(* IEC 61131-3 sources: brew/plc/plc-cellar, 2 files *)

(* ---- plc-cellar-plant.st ---- *)
(*
  plc-cellar: CherryMountain Brewery cellar PLC, full and lite variants
  (DESIGN.md 6.3, 6.7, 12.1). The ci slice runs plc-cellar.st instead.

  Per fermenter FV-101 .. FV-104:
    - on/off glycol valve control with a 0.5 degF hysteresis half band on the
      side and cone zones (cooling only)
    - the spunding setpoint: 1 psig while the beer is fermenting, 12 psig once
      the apparent extract falls below 5 degP (near terminal gravity), written
      to the RIO as absolute pressure every scan
    - the fermentation profile (FermentProfile): while CEL.PROFILE.HSnn.AUTO is
      set, the program writes both temperature setpoints for the beer's stage,
      66 degF fermenting, 70 degF for the diacetyl rest, 34 degF for the crash
      (CEL.PROFILE.TC01 to TC03, the operator's), and shows the stage in
      KSnn.STAGE. The rest lasts KC01 minutes: 180, which is 144 h of
      fermentation on the range's 48x clock. With AUTO clear the setpoints are
      the operator's. A crash raises the fermenter's temperature deviation
      alarms until the beer is cold.
  Per bright tank BBT-201 and BBT-202:
    - jacket glycol valve on/off control
    - the equilibrium head pressure for the carbonation target at the
      temperature setpoint (Zahm-Nagel fit, sea-level gauge plus 14.7 psi =
      absolute; the setpoint, not the measured temperature, so the limit does
      not swing with the glycol hysteresis), and carbonation-stone flow
      proportional to the shortfall in dissolved CO2, closed while the head is
      more than HEAD_MARGIN above that pressure or at HEAD_MAX (0.5 psi under
      the 26.1 psia high-pressure alarm), so neither that alarm nor the 15 psig
      relief valve trips in normal running. A target whose equilibrium is above
      HEAD_MAX - HEAD_MARGIN cannot be reached, so AT01.SP is clamped to the
      most that can (VOL_MAX, solved from the same fit), and the HMI shows it.
    - BBT-202 feeds the bottling line: its outlet opens while it holds beer
  Shared equipment:
    - the cellar CO2 life-safety interlock (DESIGN.md 6.7): CEL.SYS.XS01.CO2_OK
      is the hardwired, de-energize-to-trip relay from bas-vent. While it is
      open, and for CO2_RELEASE_DELAY after it closes again, the program sets
      CO2_INHIBIT, closes both carbonation valves, and closes the hop-port CO2
      purge (holding a dry-hop sequence in its purge step). No supervisory host
      takes part. The relay reads open until the building federate first
      reports it, so carbonation starts inhibited.
    - the dry-hop sequence on an operator request: CO2 purge, then dose
    - the transfer and CIP peer status bits that plc-utilities reads
    - confined-space entry (29 CFR 1910.146, DESIGN.md 6.3): a vessel's entry
      permit bit locks out its glycol valves, the bright tanks' carbonation
      stone and outlet, and (through plc-utilities) its CIP circuit, vents a
      fermenter's head through its spunding valve, holds the dry-hop doser
      while any fermenter is entered, and latches a critical alarm when a
      locked-out output is found written between scans
  Alarms (every bit in alarms.json for this PLC) are generated by
  plc/common/plcbuild.py at the ALARMS marker, with their deadbands and delays.

  Units: analog values are raw registers, engineering value x 10^scaling
  (degF x 100, psia x 100, vol x 100, % x 10). Setpoints in %MW belong to the
  operator after the first scan; the program loads defaults once and clamps.
*)

(* One glycol zone: cooling-only on/off valve with hysteresis. *)
FUNCTION_BLOCK GlycolZone
  VAR_INPUT
    PV : UINT;                 (* temperature, degF x 100 *)
    SP : UINT;                 (* setpoint, degF x 100 *)
    HYST : UINT := 50;         (* half band, 0.5 degF *)
  END_VAR
  VAR_OUTPUT
    VALVE : BOOL;              (* TRUE = open (cooling) *)
  END_VAR
  IF PV >= SP + HYST THEN
    VALVE := TRUE;
  ELSIF PV + HYST <= SP THEN
    VALVE := FALSE;
  END_IF;
END_FUNCTION_BLOCK

(* Carbonation for one bright tank. *)
FUNCTION_BLOCK Carbonation
  VAR_INPUT
    TEMP_SP : UINT;            (* temperature setpoint, degF x 100 *)
    VOL_SP : UINT;             (* target, vol x 100 *)
    VOL_PV : UINT;             (* inline meter, vol x 100 *)
    PSIA_PV : UINT;            (* head pressure, psia x 100 *)
    INHIBIT : BOOL;            (* cellar CO2 interlock *)
    HEAD_MARGIN : UINT := 50;  (* stone closes 0.5 psi above equilibrium, psi x 100 *)
    HEAD_MAX : UINT := 2560;   (* and never above 25.6 psia, psia x 100 *)
  END_VAR
  VAR_OUTPUT
    PSIA_SP : UINT;            (* equilibrium head pressure, psia x 100 *)
    VALVE : UINT;              (* stone flow valve, % x 10 *)
    VOL_MAX : UINT;            (* most reachable under HEAD_MAX, vol x 100 *)
  END_VAR
  VAR
    temp_f : REAL;
    vol : REAL;
    psig_sea_level : REAL;
    shortfall : REAL;
    qa : REAL;
    qb : REAL;
    qc : REAL;
  END_VAR
  temp_f := UINT_TO_REAL(TEMP_SP) / 100.0;
  (* The fit is quadratic in vol: qa vol^2 + qb vol + qc = 0 at the highest
     equilibrium the stone may build to (HEAD_MAX - HEAD_MARGIN). *)
  qa := -0.0684226;
  qb := 4.24267 + 0.173354 * temp_f;
  qc := -16.6999 - 0.0101059 * temp_f + 0.00116512 * temp_f * temp_f
    - (UINT_TO_REAL(HEAD_MAX - HEAD_MARGIN) / 100.0 - 14.7);
  VOL_MAX := REAL_TO_UINT(LIMIT(0.0,
    (SQRT(qb * qb - 4.0 * qa * qc) - qb) / (2.0 * qa) * 100.0, 500.0));
  vol := UINT_TO_REAL(MIN(VOL_SP, VOL_MAX)) / 100.0;
  psig_sea_level := -16.6999 - 0.0101059 * temp_f + 0.00116512 * temp_f * temp_f
    + 0.173354 * temp_f * vol + 4.24267 * vol - 0.0684226 * vol * vol;
  PSIA_SP := REAL_TO_UINT(LIMIT(0.0, (psig_sea_level + 14.7) * 100.0, 4000.0));
  (* 100 % at 0.5 vol or more short of the target, closed at the target. *)
  shortfall := vol - UINT_TO_REAL(VOL_PV) / 100.0;
  IF INHIBIT OR shortfall <= 0.0 OR PSIA_PV >= MIN(PSIA_SP + HEAD_MARGIN, HEAD_MAX) THEN
    VALVE := 0;
  ELSE
    VALVE := REAL_TO_UINT(LIMIT(0.0, shortfall * 2000.0, 1000.0));
  END_IF;
END_FUNCTION_BLOCK

(* The fermentation profile of one fermenter (DESIGN.md 6.3): which stage the
   beer is in, and the temperature that goes with it. A stage follows from the
   density meter: a vessel that reads no extract is empty, wort above TERMINAL is
   fermenting, and beer under it rests warm for REST_MIN minutes (counted in
   scans) and is then crashed. A reading must hold for SETTLE_MS before it ends
   a stage: a meter that drops out for a scan or a few seconds has not emptied
   the vessel or finished the fermentation, and the stage it would end is one
   the program cannot get back to. Beer the program has not followed from its
   fill (after a start of the PLC) is taken as crashed when it is already cold,
   and as starting its rest otherwise.

   The setpoint is one the vessel can follow, so that the deviation alarm means
   a fault and not a stage:
   - A fermenter has jackets and no heater. On the way up (wort pitched under
     the fermentation temperature, the free rise to the rest) the setpoint
     leads the beer by LEAD and goes no higher than the stage's temperature. It
     does not come back down with the beer: beer that cools in these stages has
     a glycol valve that leaks. Only a fill is different: for FILL_MS after a
     fermentation starts the setpoint follows the vessel down too, to the
     temperature of the wort that is coming in.
   - The crash falls from where the beer is toward the glycol's temperature, by
     CRASH_PCT_H percent of what is left each hour, and stops at CRASH_SP. That
     is the curve of a jacketed tank, a little slower than this one cools, so
     beer that falls behind it has lost its cooling.
   - An empty vessel's setpoint stays LEAD above the vessel: its jackets stay
     shut, the next wort is not chilled on its way in, and nothing alarms. *)
FUNCTION_BLOCK FermentProfile
  VAR_INPUT
    EXTRACT : UINT;            (* apparent extract, degP x 100 *)
    TEMP : UINT;               (* side temperature, degF x 100 *)
    FERMENT_SP : UINT;         (* temperature while fermenting, degF x 100 *)
    REST_SP : UINT;            (* temperature of the diacetyl rest, degF x 100 *)
    CRASH_SP : UINT;           (* temperature of the crash, degF x 100 *)
    REST_MIN : UINT;           (* rest length, minutes *)
    SCAN_MS : UDINT;           (* the task interval, ms *)
    EMPTY : UINT := 50;        (* under 0.5 degP the vessel is empty *)
    TERMINAL : UINT := 500;    (* under 5 degP the beer is near terminal gravity *)
    COLD : UINT := 6000;       (* under 60 degF the beer has been crashed *)
    SETTLE_MS : UDINT := 60000;  (* a reading ends a stage once it has held this long *)
    LEAD : UINT := 100;        (* on the way up the setpoint leads the beer by 1 degF *)
    GLYCOL : UINT := 2800;     (* the glycol supply, degF x 100: the crash falls toward it *)
    CRASH_PCT_H : UINT := 25;  (* ... by this share of what is left, each hour *)
    SP_MIN : UINT := 2000;     (* the setpoint limits of the program *)
    SP_MAX : UINT := 9000;
    FILL_MS : UDINT := 1800000;  (* a knockout into the vessel is over in this time *)
  END_VAR
  VAR_OUTPUT
    STAGE : UINT;              (* 0 empty, 1 fermenting, 2 diacetyl rest, 3 crash *)
    SP : UINT;                 (* the stage's setpoint now, degF x 100 *)
  END_VAR
  VAR
    rest_ms : UDINT;           (* time in the rest so far *)
    empty_ms : UDINT;          (* how long the meter has read no extract *)
    terminal_ms : UDINT;       (* how long it has read under TERMINAL *)
    last_stage : UINT := 99;   (* the stage of the scan before; 99 before the first *)
    sp_now : REAL := 0.0;      (* the setpoint, degF x 100, between scans *)
    lead_sp : REAL;
    cap : REAL;
    stage_ms : UDINT;          (* time in the stage, up to FILL_MS *)
  END_VAR
  IF EXTRACT < EMPTY THEN
    empty_ms := MIN(empty_ms + SCAN_MS, SETTLE_MS);
  ELSE
    empty_ms := 0;
  END_IF;
  IF EXTRACT < TERMINAL THEN
    terminal_ms := MIN(terminal_ms + SCAN_MS, SETTLE_MS);
  ELSE
    terminal_ms := 0;
  END_IF;
  IF EXTRACT < EMPTY THEN
    (* Until the reading has held, the stage stays as it is (and a rest's clock
       waits): this may be the meter, not the vessel. *)
    IF empty_ms >= SETTLE_MS THEN
      STAGE := 0;
    END_IF;
  ELSIF STAGE = 0 THEN
    IF EXTRACT >= TERMINAL THEN
      STAGE := 1;
    ELSIF TEMP < COLD THEN
      STAGE := 3;
    ELSE
      STAGE := 2;
      rest_ms := 0;
    END_IF;
  ELSIF STAGE = 1 THEN
    IF terminal_ms >= SETTLE_MS THEN
      STAGE := 2;
      rest_ms := 0;
    END_IF;
  ELSIF STAGE = 2 THEN
    IF rest_ms >= UINT_TO_UDINT(REST_MIN) * 60000 THEN
      STAGE := 3;
    ELSE
      rest_ms := rest_ms + SCAN_MS;
    END_IF;
  END_IF;

  lead_sp := UINT_TO_REAL(TEMP) + UINT_TO_REAL(LEAD);
  IF STAGE = 3 THEN
    IF last_stage <> 3 THEN
      sp_now := UINT_TO_REAL(TEMP);   (* the crash starts from where the beer is *)
    END_IF;
    sp_now := sp_now - (sp_now - UINT_TO_REAL(GLYCOL)) * UINT_TO_REAL(CRASH_PCT_H) / 100.0
      * UDINT_TO_REAL(SCAN_MS) / 3600000.0;
    sp_now := MAX(sp_now, UINT_TO_REAL(CRASH_SP));
  ELSIF STAGE = 0 THEN
    sp_now := lead_sp;
  ELSE
    IF STAGE = 2 THEN
      cap := UINT_TO_REAL(REST_SP);
    ELSE
      cap := UINT_TO_REAL(FERMENT_SP);
    END_IF;
    IF last_stage <> STAGE THEN
      stage_ms := 0;
      IF last_stage <> 1 THEN
        sp_now := 0.0;                (* nothing to carry over: start from the beer *)
      END_IF;
    ELSE
      stage_ms := MIN(stage_ms + SCAN_MS, FILL_MS);
    END_IF;
    IF STAGE = 1 AND stage_ms < FILL_MS THEN
      sp_now := MIN(cap, lead_sp);    (* a fill: down to the wort's temperature too *)
    ELSE
      sp_now := MIN(cap, MAX(sp_now, lead_sp));
    END_IF;
  END_IF;
  last_stage := STAGE;
  SP := REAL_TO_UINT(LIMIT(UINT_TO_REAL(SP_MIN), sp_now, UINT_TO_REAL(SP_MAX)));
END_FUNCTION_BLOCK

PROGRAM plc_cellar
  (* LOCATED_VARS: plcbuild.py splices the located variables and alarm instances here. *)

  VAR CONSTANT
    TEMP_SP_MIN : UINT := 2000;       (* 20 degF *)
    TEMP_SP_MAX : UINT := 9000;       (* 90 degF *)
    VOL_SP_MAX : UINT := 350;         (* 3.5 vol *)
    AMBIENT_PSIA : UINT := 1210;      (* 12.1 psia at 5,200 ft *)
    SPUND_LOW_PSIG : UINT := 100;     (* 1 psig while fermenting *)
    SPUND_HIGH_PSIG : UINT := 1200;   (* 12 psig near terminal gravity *)
    TERMINAL_PLATO : UINT := 500;     (* 5 degP *)
    BBT_FEED_MIN_LEVEL : UINT := 50;  (* 5 % *)
    CO2_RELEASE_DELAY : TIME := T#60s;  (* relay must be healthy this long *)
    DH_PURGE_TIME : TIME := T#30s;      (* hop-port CO2 purge before a dose *)
    DH_DOSE_TIME : TIME := T#60s;       (* dose valve open *)
    SCAN_MS : UDINT := 100;           (* the task interval plcbuild.py sets (T#100ms) *)
    REST_MIN_MAX : UINT := 6000;      (* 100 h *)
  END_VAR

  VAR
    started : BOOL := FALSE;
    fv101_side : GlycolZone;
    fv101_cone : GlycolZone;
    fv102_side : GlycolZone;
    fv102_cone : GlycolZone;
    fv103_side : GlycolZone;
    fv103_cone : GlycolZone;
    fv104_side : GlycolZone;
    fv104_cone : GlycolZone;
    fv101_profile : FermentProfile;
    fv102_profile : FermentProfile;
    fv103_profile : FermentProfile;
    fv104_profile : FermentProfile;
    bbt201_zone : GlycolZone;
    bbt202_zone : GlycolZone;
    bbt201_carb : Carbonation;
    bbt202_carb : Carbonation;
    co2_healthy : TON;
    transfer_active : BOOL;
    dh_step : INT := 0;
    dh_purge : TON;
    dh_dose : TON;
    fv_entry : BOOL;
  END_VAR

  (* First scan: default setpoints for the staggered initial state (DESIGN.md 9.4). *)
  IF NOT started THEN
    CEL_FV101_TT01_SP := 6600;
    CEL_FV101_TT02_SP := 6600;
    CEL_FV102_TT01_SP := 6600;
    CEL_FV102_TT02_SP := 6600;
    CEL_FV103_TT01_SP := 6800;
    CEL_FV103_TT02_SP := 6800;
    CEL_FV104_TT01_SP := 3400;
    CEL_FV104_TT02_SP := 3400;
    CEL_BBT201_TT01_SP := 3400;
    CEL_BBT202_TT01_SP := 3400;
    CEL_BBT201_AT01_SP := 260;
    CEL_BBT202_AT01_SP := 260;
    (* The recipe's profile (fire-of-the-phenix), on for every fermenter. *)
    CEL_PROFILE_TC01_SP := 6600;
    CEL_PROFILE_TC02_SP := 7000;
    CEL_PROFILE_TC03_SP := 3400;
    CEL_PROFILE_KC01_SP := 180;
    CEL_PROFILE_HS01_AUTO := TRUE;
    CEL_PROFILE_HS02_AUTO := TRUE;
    CEL_PROFILE_HS03_AUTO := TRUE;
    CEL_PROFILE_HS04_AUTO := TRUE;
    started := TRUE;
  END_IF;

  CEL_FV101_TT01_SP := LIMIT(TEMP_SP_MIN, CEL_FV101_TT01_SP, TEMP_SP_MAX);
  CEL_FV101_TT02_SP := LIMIT(TEMP_SP_MIN, CEL_FV101_TT02_SP, TEMP_SP_MAX);
  CEL_FV102_TT01_SP := LIMIT(TEMP_SP_MIN, CEL_FV102_TT01_SP, TEMP_SP_MAX);
  CEL_FV102_TT02_SP := LIMIT(TEMP_SP_MIN, CEL_FV102_TT02_SP, TEMP_SP_MAX);
  CEL_FV103_TT01_SP := LIMIT(TEMP_SP_MIN, CEL_FV103_TT01_SP, TEMP_SP_MAX);
  CEL_FV103_TT02_SP := LIMIT(TEMP_SP_MIN, CEL_FV103_TT02_SP, TEMP_SP_MAX);
  CEL_FV104_TT01_SP := LIMIT(TEMP_SP_MIN, CEL_FV104_TT01_SP, TEMP_SP_MAX);
  CEL_FV104_TT02_SP := LIMIT(TEMP_SP_MIN, CEL_FV104_TT02_SP, TEMP_SP_MAX);
  CEL_BBT201_TT01_SP := LIMIT(TEMP_SP_MIN, CEL_BBT201_TT01_SP, TEMP_SP_MAX);
  CEL_BBT202_TT01_SP := LIMIT(TEMP_SP_MIN, CEL_BBT202_TT01_SP, TEMP_SP_MAX);
  CEL_BBT201_AT01_SP := MIN(CEL_BBT201_AT01_SP, VOL_SP_MAX);
  CEL_BBT202_AT01_SP := MIN(CEL_BBT202_AT01_SP, VOL_SP_MAX);
  CEL_PROFILE_TC01_SP := LIMIT(TEMP_SP_MIN, CEL_PROFILE_TC01_SP, TEMP_SP_MAX);
  CEL_PROFILE_TC02_SP := LIMIT(TEMP_SP_MIN, CEL_PROFILE_TC02_SP, TEMP_SP_MAX);
  CEL_PROFILE_TC03_SP := LIMIT(TEMP_SP_MIN, CEL_PROFILE_TC03_SP, TEMP_SP_MAX);
  CEL_PROFILE_KC01_SP := MIN(CEL_PROFILE_KC01_SP, REST_MIN_MAX);

  (* ---- fermentation profile: the stage's temperature for a fermenter on AUTO --- *)
  fv101_profile(EXTRACT := CEL_FV101_DT01_PV, TEMP := CEL_FV101_TT01_PV,
    FERMENT_SP := CEL_PROFILE_TC01_SP, REST_SP := CEL_PROFILE_TC02_SP,
    CRASH_SP := CEL_PROFILE_TC03_SP, REST_MIN := CEL_PROFILE_KC01_SP, SCAN_MS := SCAN_MS);
  CEL_PROFILE_KS01_STAGE := fv101_profile.STAGE;
  IF CEL_PROFILE_HS01_AUTO THEN
    CEL_FV101_TT01_SP := fv101_profile.SP;
    CEL_FV101_TT02_SP := fv101_profile.SP;
  END_IF;
  fv102_profile(EXTRACT := CEL_FV102_DT01_PV, TEMP := CEL_FV102_TT01_PV,
    FERMENT_SP := CEL_PROFILE_TC01_SP, REST_SP := CEL_PROFILE_TC02_SP,
    CRASH_SP := CEL_PROFILE_TC03_SP, REST_MIN := CEL_PROFILE_KC01_SP, SCAN_MS := SCAN_MS);
  CEL_PROFILE_KS02_STAGE := fv102_profile.STAGE;
  IF CEL_PROFILE_HS02_AUTO THEN
    CEL_FV102_TT01_SP := fv102_profile.SP;
    CEL_FV102_TT02_SP := fv102_profile.SP;
  END_IF;
  fv103_profile(EXTRACT := CEL_FV103_DT01_PV, TEMP := CEL_FV103_TT01_PV,
    FERMENT_SP := CEL_PROFILE_TC01_SP, REST_SP := CEL_PROFILE_TC02_SP,
    CRASH_SP := CEL_PROFILE_TC03_SP, REST_MIN := CEL_PROFILE_KC01_SP, SCAN_MS := SCAN_MS);
  CEL_PROFILE_KS03_STAGE := fv103_profile.STAGE;
  IF CEL_PROFILE_HS03_AUTO THEN
    CEL_FV103_TT01_SP := fv103_profile.SP;
    CEL_FV103_TT02_SP := fv103_profile.SP;
  END_IF;
  fv104_profile(EXTRACT := CEL_FV104_DT01_PV, TEMP := CEL_FV104_TT01_PV,
    FERMENT_SP := CEL_PROFILE_TC01_SP, REST_SP := CEL_PROFILE_TC02_SP,
    CRASH_SP := CEL_PROFILE_TC03_SP, REST_MIN := CEL_PROFILE_KC01_SP, SCAN_MS := SCAN_MS);
  CEL_PROFILE_KS04_STAGE := fv104_profile.STAGE;
  IF CEL_PROFILE_HS04_AUTO THEN
    CEL_FV104_TT01_SP := fv104_profile.SP;
    CEL_FV104_TT02_SP := fv104_profile.SP;
  END_IF;

  (* ---- confined-space entry (29 CFR 1910.146, DESIGN.md 6.3) ------------------ *)
  (* The entry supervisor sets HSnn.ENTRY when the permit is issued. The program
     leaves every locked-out output off at the end of a scan, so a locked output
     that is on at the top of this one was written in between (an HMI, the EWS,
     or an attacker on the PLC's Modbus server): XAnn latches until the entry
     ends. *)
  CEL_ENTRY_XA01_PV := CEL_ENTRY_XS01_LOCKED
    AND (CEL_ENTRY_XA01_PV OR CEL_FV101_TV01_CMD OR CEL_FV101_TV02_CMD);
  CEL_ENTRY_XA02_PV := CEL_ENTRY_XS02_LOCKED
    AND (CEL_ENTRY_XA02_PV OR CEL_FV102_TV01_CMD OR CEL_FV102_TV02_CMD);
  CEL_ENTRY_XA03_PV := CEL_ENTRY_XS03_LOCKED
    AND (CEL_ENTRY_XA03_PV OR CEL_FV103_TV01_CMD OR CEL_FV103_TV02_CMD);
  CEL_ENTRY_XA04_PV := CEL_ENTRY_XS04_LOCKED
    AND (CEL_ENTRY_XA04_PV OR CEL_FV104_TV01_CMD OR CEL_FV104_TV02_CMD);
  CEL_ENTRY_XA05_PV := CEL_ENTRY_XS05_LOCKED
    AND (CEL_ENTRY_XA05_PV OR CEL_BBT201_TV01_CMD OR CEL_BBT201_XV01_CMD OR CEL_BBT201_FCV01_OUT > 0);
  CEL_ENTRY_XA06_PV := CEL_ENTRY_XS06_LOCKED
    AND (CEL_ENTRY_XA06_PV OR CEL_BBT202_TV01_CMD OR CEL_BBT202_XV01_CMD OR CEL_BBT202_FCV01_OUT > 0);
  CEL_ENTRY_XS01_LOCKED := CEL_ENTRY_HS01_ENTRY;
  CEL_ENTRY_XS11_CIP_OK := NOT CEL_ENTRY_XS01_LOCKED;
  CEL_ENTRY_XS02_LOCKED := CEL_ENTRY_HS02_ENTRY;
  CEL_ENTRY_XS12_CIP_OK := NOT CEL_ENTRY_XS02_LOCKED;
  CEL_ENTRY_XS03_LOCKED := CEL_ENTRY_HS03_ENTRY;
  CEL_ENTRY_XS13_CIP_OK := NOT CEL_ENTRY_XS03_LOCKED;
  CEL_ENTRY_XS04_LOCKED := CEL_ENTRY_HS04_ENTRY;
  CEL_ENTRY_XS14_CIP_OK := NOT CEL_ENTRY_XS04_LOCKED;
  CEL_ENTRY_XS05_LOCKED := CEL_ENTRY_HS05_ENTRY;
  CEL_ENTRY_XS15_CIP_OK := NOT CEL_ENTRY_XS05_LOCKED;
  CEL_ENTRY_XS06_LOCKED := CEL_ENTRY_HS06_ENTRY;
  CEL_ENTRY_XS16_CIP_OK := NOT CEL_ENTRY_XS06_LOCKED;
  fv_entry := CEL_ENTRY_XS01_LOCKED OR CEL_ENTRY_XS02_LOCKED
    OR CEL_ENTRY_XS03_LOCKED OR CEL_ENTRY_XS04_LOCKED;

  (* ---- CO2 life-safety interlock (DESIGN.md 6.7) ---------------------------- *)
  (* The relay is de-energize to trip: open (FALSE) inhibits at once, and the
     inhibit clears only after the relay has been healthy for CO2_RELEASE_DELAY. *)
  co2_healthy(IN := CEL_SYS_XS01_CO2_OK, PT := CO2_RELEASE_DELAY);
  CEL_SYS_XS01_CO2_INHIBIT := NOT co2_healthy.Q;

  (* ---- fermenters --------------------------------------------------------------- *)
  fv101_side(PV := CEL_FV101_TT01_PV, SP := CEL_FV101_TT01_SP);
  CEL_FV101_TV01_CMD := fv101_side.VALVE;
  fv101_cone(PV := CEL_FV101_TT02_PV, SP := CEL_FV101_TT02_SP);
  CEL_FV101_TV02_CMD := fv101_cone.VALVE;
  IF CEL_FV101_DT01_PV < TERMINAL_PLATO THEN
    CEL_FV101_PCV01_SP := SPUND_HIGH_PSIG + AMBIENT_PSIA;
  ELSE
    CEL_FV101_PCV01_SP := SPUND_LOW_PSIG + AMBIENT_PSIA;
  END_IF;

  fv102_side(PV := CEL_FV102_TT01_PV, SP := CEL_FV102_TT01_SP);
  CEL_FV102_TV01_CMD := fv102_side.VALVE;
  fv102_cone(PV := CEL_FV102_TT02_PV, SP := CEL_FV102_TT02_SP);
  CEL_FV102_TV02_CMD := fv102_cone.VALVE;
  IF CEL_FV102_DT01_PV < TERMINAL_PLATO THEN
    CEL_FV102_PCV01_SP := SPUND_HIGH_PSIG + AMBIENT_PSIA;
  ELSE
    CEL_FV102_PCV01_SP := SPUND_LOW_PSIG + AMBIENT_PSIA;
  END_IF;

  fv103_side(PV := CEL_FV103_TT01_PV, SP := CEL_FV103_TT01_SP);
  CEL_FV103_TV01_CMD := fv103_side.VALVE;
  fv103_cone(PV := CEL_FV103_TT02_PV, SP := CEL_FV103_TT02_SP);
  CEL_FV103_TV02_CMD := fv103_cone.VALVE;
  IF CEL_FV103_DT01_PV < TERMINAL_PLATO THEN
    CEL_FV103_PCV01_SP := SPUND_HIGH_PSIG + AMBIENT_PSIA;
  ELSE
    CEL_FV103_PCV01_SP := SPUND_LOW_PSIG + AMBIENT_PSIA;
  END_IF;

  fv104_side(PV := CEL_FV104_TT01_PV, SP := CEL_FV104_TT01_SP);
  CEL_FV104_TV01_CMD := fv104_side.VALVE;
  fv104_cone(PV := CEL_FV104_TT02_PV, SP := CEL_FV104_TT02_SP);
  CEL_FV104_TV02_CMD := fv104_cone.VALVE;
  IF CEL_FV104_DT01_PV < TERMINAL_PLATO THEN
    CEL_FV104_PCV01_SP := SPUND_HIGH_PSIG + AMBIENT_PSIA;
  ELSE
    CEL_FV104_PCV01_SP := SPUND_LOW_PSIG + AMBIENT_PSIA;
  END_IF;

  (* ---- bright tanks --------------------------------------------------------------- *)
  bbt201_zone(PV := CEL_BBT201_TT01_PV, SP := CEL_BBT201_TT01_SP);
  CEL_BBT201_TV01_CMD := bbt201_zone.VALVE;
  bbt201_carb(TEMP_SP := CEL_BBT201_TT01_SP, VOL_SP := CEL_BBT201_AT01_SP,
    VOL_PV := CEL_BBT201_AT01_PV, PSIA_PV := CEL_BBT201_PT01_PV,
    INHIBIT := CEL_SYS_XS01_CO2_INHIBIT);
  CEL_BBT201_PT01_SP := bbt201_carb.PSIA_SP;
  CEL_BBT201_AT01_SP := MIN(CEL_BBT201_AT01_SP, bbt201_carb.VOL_MAX);
  CEL_BBT201_FCV01_OUT := bbt201_carb.VALVE;
  CEL_BBT201_XV01_CMD := FALSE;  (* BBT-201 is carbonating, not feeding *)

  bbt202_zone(PV := CEL_BBT202_TT01_PV, SP := CEL_BBT202_TT01_SP);
  CEL_BBT202_TV01_CMD := bbt202_zone.VALVE;
  bbt202_carb(TEMP_SP := CEL_BBT202_TT01_SP, VOL_SP := CEL_BBT202_AT01_SP,
    VOL_PV := CEL_BBT202_AT01_PV, PSIA_PV := CEL_BBT202_PT01_PV,
    INHIBIT := CEL_SYS_XS01_CO2_INHIBIT);
  CEL_BBT202_PT01_SP := bbt202_carb.PSIA_SP;
  CEL_BBT202_AT01_SP := MIN(CEL_BBT202_AT01_SP, bbt202_carb.VOL_MAX);
  CEL_BBT202_FCV01_OUT := bbt202_carb.VALVE;
  CEL_BBT202_XV01_CMD := CEL_BBT202_LT01_PV > BBT_FEED_MIN_LEVEL;

  (* ---- entry lockout: glycol, carbonation CO2, and outlet off; the fermenter's
     head vented through its spunding valve (setpoint at ambient, 0 psig). -- *)
  IF CEL_ENTRY_XS01_LOCKED THEN
    CEL_FV101_TV01_CMD := FALSE;
    CEL_FV101_TV02_CMD := FALSE;
    CEL_FV101_PCV01_SP := AMBIENT_PSIA;
  END_IF;
  IF CEL_ENTRY_XS02_LOCKED THEN
    CEL_FV102_TV01_CMD := FALSE;
    CEL_FV102_TV02_CMD := FALSE;
    CEL_FV102_PCV01_SP := AMBIENT_PSIA;
  END_IF;
  IF CEL_ENTRY_XS03_LOCKED THEN
    CEL_FV103_TV01_CMD := FALSE;
    CEL_FV103_TV02_CMD := FALSE;
    CEL_FV103_PCV01_SP := AMBIENT_PSIA;
  END_IF;
  IF CEL_ENTRY_XS04_LOCKED THEN
    CEL_FV104_TV01_CMD := FALSE;
    CEL_FV104_TV02_CMD := FALSE;
    CEL_FV104_PCV01_SP := AMBIENT_PSIA;
  END_IF;
  IF CEL_ENTRY_XS05_LOCKED THEN
    CEL_BBT201_TV01_CMD := FALSE;
    CEL_BBT201_XV01_CMD := FALSE;
    CEL_BBT201_FCV01_OUT := 0;
  END_IF;
  IF CEL_ENTRY_XS06_LOCKED THEN
    CEL_BBT202_TV01_CMD := FALSE;
    CEL_BBT202_XV01_CMD := FALSE;
    CEL_BBT202_FCV01_OUT := 0;
  END_IF;

  (* ---- dry-hop doser (DESIGN.md 6.3): the operator sets the dose request
     (CEL.DH.XC01.CMD); the PLC purges the hop port with CO2 for DH_PURGE_TIME,
     doses for DH_DOSE_TIME, and clears the request. The CO2 interlock closes the
     purge and holds the sequence (the purge timer restarts) while it is set, so
     no CO2 goes into a cellar that is already at tier 2 (DESIGN.md 6.7). *)
  CASE dh_step OF
    0:
      IF CEL_DH_XC01_CMD AND NOT fv_entry THEN
        dh_step := 1;
      END_IF;
    1:
      IF NOT CEL_DH_XC01_CMD THEN
        dh_step := 0;  (* the operator withdrew the request *)
      ELSIF dh_purge.Q THEN
        dh_step := 2;
      END_IF;
    2:
      IF dh_dose.Q THEN
        dh_step := 0;
        CEL_DH_XC01_CMD := FALSE;
      END_IF;
  ELSE
    dh_step := 0;
  END_CASE;
  CEL_DH_XV01_CMD := (dh_step = 1) AND NOT CEL_SYS_XS01_CO2_INHIBIT AND NOT fv_entry;
  dh_purge(IN := CEL_DH_XV01_CMD, PT := DH_PURGE_TIME);
  CEL_DH_XV02_CMD := dh_step = 2 AND NOT fv_entry;
  dh_dose(IN := CEL_DH_XV02_CMD, PT := DH_DOSE_TIME);
  CEL_DH_XS01_STEP := INT_TO_UINT(dh_step);

  (* ---- transfer panel and the peer status for plc-utilities (DESIGN.md 6.6 #4) *)
  CEL_XFER_HS01_CMD := FALSE;
  transfer_active := CEL_XFER_YS01_PV OR CEL_XFER_HS01_CMD;
  CEL_XFER_XS01_ACTIVE := transfer_active;
  CEL_XFER_XS02_CIP_PERMIT := NOT transfer_active;

  (* ALARMS: plcbuild.py generates the alarm logic here. *)
END_PROGRAM

(* ---- plc-cellar.st ---- *)
(*
  plc-cellar: CherryMountain Brewery cellar PLC (ci variant, DESIGN.md 12.1).

  Per fermenter FV-101 .. FV-104 this program runs:
    - on/off glycol valve control with hysteresis on the side and cone zones
    - a spunding valve pressure setpoint, written to the RIO every scan
    - ISA-18.2 alarm evaluation with on-delay timers (limits and delays below
      come from plant/generated/ci/alarms.json; assemble.py checks they match)

  Units: every analog value is a raw unsigned register, engineering value x 100
  (degF for temperatures, psia for pressures). Setpoints in %MW are written by
  the operator (FUXA, Modbus holding registers from qw_count, see
  modbus_slave.json); the PLC loads defaults once at start-up and clamps them
  to the plant range afterwards.

  The located variables (the %IW/%QX/%QW/%MW map) are not written here. They
  come from plant/generated/ci/openplc/plc-cellar/located_vars.st, and
  assemble.py splices that VAR block in at the marker comment in plc_cellar.
  Do not hand-edit addresses: change plant/plant.yaml and rerun plantgen.
*)

(* One glycol zone: on/off valve with hysteresis plus its temperature alarms. *)
FUNCTION_BLOCK ZoneControl
  VAR_INPUT
    PV : UINT;                 (* temperature, degF x 100 *)
    SP : UINT;                 (* setpoint, degF x 100 *)
    HYST : UINT := 50;         (* valve hysteresis half band, 0.5 degF *)
    DEV_LIMIT : UINT;          (* deviation alarm limit, degF x 100 *)
    DEV_DELAY : TIME;          (* deviation alarm on-delay *)
    HIGH_LIMIT : UINT;         (* high alarm limit, degF x 100; 0 = no high alarm *)
    HIGH_DELAY : TIME;         (* high alarm on-delay *)
  END_VAR
  VAR_OUTPUT
    VALVE : BOOL;              (* glycol valve command, TRUE = open (cooling) *)
    ALM_DEV : BOOL;
    ALM_HIGH : BOOL;
  END_VAR
  VAR
    dev_timer : TON;
    high_timer : TON;
    err : DINT;
    dev_cond : BOOL;
    high_cond : BOOL;
  END_VAR

  (* Cooling only: open above SP + HYST, close below SP - HYST, hold between. *)
  IF PV >= SP + HYST THEN
    VALVE := TRUE;
  ELSIF PV + HYST <= SP THEN
    VALVE := FALSE;
  END_IF;

  err := UINT_TO_DINT(PV) - UINT_TO_DINT(SP);
  dev_cond := ABS(err) > UINT_TO_DINT(DEV_LIMIT);
  dev_timer(IN := dev_cond, PT := DEV_DELAY);
  ALM_DEV := dev_timer.Q;

  high_cond := (HIGH_LIMIT > 0) AND (PV > HIGH_LIMIT);
  high_timer(IN := high_cond, PT := HIGH_DELAY);
  ALM_HIGH := high_timer.Q;
END_FUNCTION_BLOCK

(* Head pressure (absolute) high and low alarms for one fermenter. *)
FUNCTION_BLOCK PressureAlarm
  VAR_INPUT
    PV : UINT;                 (* psia x 100 *)
    HIGH_LIMIT : UINT;
    HIGH_DELAY : TIME;
    LOW_LIMIT : UINT;
    LOW_DELAY : TIME;
  END_VAR
  VAR_OUTPUT
    ALM_HIGH : BOOL;
    ALM_LOW : BOOL;
  END_VAR
  VAR
    high_timer : TON;
    low_timer : TON;
  END_VAR

  high_timer(IN := PV > HIGH_LIMIT, PT := HIGH_DELAY);
  ALM_HIGH := high_timer.Q;
  low_timer(IN := PV < LOW_LIMIT, PT := LOW_DELAY);
  ALM_LOW := low_timer.Q;
END_FUNCTION_BLOCK

PROGRAM plc_cellar
  (* LOCATED_VARS: assemble.py splices located_vars.st here. *)

  VAR CONSTANT
    (* Alarm limits and delays: keep equal to plant/generated/ci/alarms.json. *)
    TEMP_DEV_LIMIT : UINT := 200;       (* 2.0 degF *)
    TEMP_DEV_DELAY_SIDE : TIME := T#900s;
    TEMP_DEV_DELAY_CONE : TIME := T#900s;
    TEMP_HIGH_LIMIT : UINT := 7500;     (* 75.0 degF, side zone only *)
    TEMP_HIGH_DELAY : TIME := T#300s;
    PRESS_HIGH_LIMIT : UINT := 2610;    (* 26.1 psia *)
    PRESS_HIGH_DELAY : TIME := T#30s;
    PRESS_LOW_LIMIT : UINT := 1160;     (* 11.6 psia *)
    PRESS_LOW_DELAY : TIME := T#300s;
    (* Operator setpoint range, from plant.yaml (20 .. 90 degF). *)
    TEMP_SP_MIN : UINT := 2000;
    TEMP_SP_MAX : UINT := 9000;
    (* Site ambient pressure, 12.1 psia (5200 ft). *)
    AMBIENT_PSIA : UINT := 1210;
  END_VAR

  VAR
    started : BOOL := FALSE;
    (* Spunding setpoints, psig x 100. They follow the ci initial state in
       plant.yaml: FV-101/102 early fermentation, FV-103/104 sealed. *)
    spund_fv101_psig : UINT := 100;
    spund_fv102_psig : UINT := 100;
    spund_fv103_psig : UINT := 1200;
    spund_fv104_psig : UINT := 1200;

    fv101_side : ZoneControl;
    fv101_cone : ZoneControl;
    fv101_press : PressureAlarm;
    fv102_side : ZoneControl;
    fv102_cone : ZoneControl;
    fv102_press : PressureAlarm;
    fv103_side : ZoneControl;
    fv103_cone : ZoneControl;
    fv103_press : PressureAlarm;
    fv104_side : ZoneControl;
    fv104_cone : ZoneControl;
    fv104_press : PressureAlarm;
  END_VAR

  (* First scan: load default setpoints (the ci plant starts mid-fermentation). *)
  IF NOT started THEN
    CEL_FV101_TT01_SP := 6600;
    CEL_FV101_TT02_SP := 6600;
    CEL_FV102_TT01_SP := 6600;
    CEL_FV102_TT02_SP := 6600;
    CEL_FV103_TT01_SP := 6800;
    CEL_FV103_TT02_SP := 6800;
    CEL_FV104_TT01_SP := 5000;
    CEL_FV104_TT02_SP := 5000;
    started := TRUE;
  END_IF;

  (* Keep operator-written setpoints inside the plant range. *)
  CEL_FV101_TT01_SP := LIMIT(TEMP_SP_MIN, CEL_FV101_TT01_SP, TEMP_SP_MAX);
  CEL_FV101_TT02_SP := LIMIT(TEMP_SP_MIN, CEL_FV101_TT02_SP, TEMP_SP_MAX);
  CEL_FV102_TT01_SP := LIMIT(TEMP_SP_MIN, CEL_FV102_TT01_SP, TEMP_SP_MAX);
  CEL_FV102_TT02_SP := LIMIT(TEMP_SP_MIN, CEL_FV102_TT02_SP, TEMP_SP_MAX);
  CEL_FV103_TT01_SP := LIMIT(TEMP_SP_MIN, CEL_FV103_TT01_SP, TEMP_SP_MAX);
  CEL_FV103_TT02_SP := LIMIT(TEMP_SP_MIN, CEL_FV103_TT02_SP, TEMP_SP_MAX);
  CEL_FV104_TT01_SP := LIMIT(TEMP_SP_MIN, CEL_FV104_TT01_SP, TEMP_SP_MAX);
  CEL_FV104_TT02_SP := LIMIT(TEMP_SP_MIN, CEL_FV104_TT02_SP, TEMP_SP_MAX);

  (* FV-101 *)
  fv101_side(PV := CEL_FV101_TT01_PV, SP := CEL_FV101_TT01_SP,
    DEV_LIMIT := TEMP_DEV_LIMIT, DEV_DELAY := TEMP_DEV_DELAY_SIDE,
    HIGH_LIMIT := TEMP_HIGH_LIMIT, HIGH_DELAY := TEMP_HIGH_DELAY);
  CEL_FV101_TV01_CMD := fv101_side.VALVE;
  CEL_FV101_TT01_ALM_DEVIATION := fv101_side.ALM_DEV;
  CEL_FV101_TT01_ALM_HIGH := fv101_side.ALM_HIGH;

  fv101_cone(PV := CEL_FV101_TT02_PV, SP := CEL_FV101_TT02_SP,
    DEV_LIMIT := TEMP_DEV_LIMIT, DEV_DELAY := TEMP_DEV_DELAY_CONE,
    HIGH_LIMIT := 0, HIGH_DELAY := T#0s);
  CEL_FV101_TV02_CMD := fv101_cone.VALVE;
  CEL_FV101_TT02_ALM_DEVIATION := fv101_cone.ALM_DEV;

  fv101_press(PV := CEL_FV101_PT01_PV,
    HIGH_LIMIT := PRESS_HIGH_LIMIT, HIGH_DELAY := PRESS_HIGH_DELAY,
    LOW_LIMIT := PRESS_LOW_LIMIT, LOW_DELAY := PRESS_LOW_DELAY);
  CEL_FV101_PT01_ALM_HIGH := fv101_press.ALM_HIGH;
  CEL_FV101_PT01_ALM_LOW := fv101_press.ALM_LOW;

  (* Spunding setpoint to the RIO, absolute psia x 100, every scan. *)
  CEL_FV101_PCV01_SP := spund_fv101_psig + AMBIENT_PSIA;

  (* FV-102 *)
  fv102_side(PV := CEL_FV102_TT01_PV, SP := CEL_FV102_TT01_SP,
    DEV_LIMIT := TEMP_DEV_LIMIT, DEV_DELAY := TEMP_DEV_DELAY_SIDE,
    HIGH_LIMIT := TEMP_HIGH_LIMIT, HIGH_DELAY := TEMP_HIGH_DELAY);
  CEL_FV102_TV01_CMD := fv102_side.VALVE;
  CEL_FV102_TT01_ALM_DEVIATION := fv102_side.ALM_DEV;
  CEL_FV102_TT01_ALM_HIGH := fv102_side.ALM_HIGH;

  fv102_cone(PV := CEL_FV102_TT02_PV, SP := CEL_FV102_TT02_SP,
    DEV_LIMIT := TEMP_DEV_LIMIT, DEV_DELAY := TEMP_DEV_DELAY_CONE,
    HIGH_LIMIT := 0, HIGH_DELAY := T#0s);
  CEL_FV102_TV02_CMD := fv102_cone.VALVE;
  CEL_FV102_TT02_ALM_DEVIATION := fv102_cone.ALM_DEV;

  fv102_press(PV := CEL_FV102_PT01_PV,
    HIGH_LIMIT := PRESS_HIGH_LIMIT, HIGH_DELAY := PRESS_HIGH_DELAY,
    LOW_LIMIT := PRESS_LOW_LIMIT, LOW_DELAY := PRESS_LOW_DELAY);
  CEL_FV102_PT01_ALM_HIGH := fv102_press.ALM_HIGH;
  CEL_FV102_PT01_ALM_LOW := fv102_press.ALM_LOW;

  (* Spunding setpoint to the RIO, absolute psia x 100, every scan. *)
  CEL_FV102_PCV01_SP := spund_fv102_psig + AMBIENT_PSIA;

  (* FV-103 *)
  fv103_side(PV := CEL_FV103_TT01_PV, SP := CEL_FV103_TT01_SP,
    DEV_LIMIT := TEMP_DEV_LIMIT, DEV_DELAY := TEMP_DEV_DELAY_SIDE,
    HIGH_LIMIT := TEMP_HIGH_LIMIT, HIGH_DELAY := TEMP_HIGH_DELAY);
  CEL_FV103_TV01_CMD := fv103_side.VALVE;
  CEL_FV103_TT01_ALM_DEVIATION := fv103_side.ALM_DEV;
  CEL_FV103_TT01_ALM_HIGH := fv103_side.ALM_HIGH;

  fv103_cone(PV := CEL_FV103_TT02_PV, SP := CEL_FV103_TT02_SP,
    DEV_LIMIT := TEMP_DEV_LIMIT, DEV_DELAY := TEMP_DEV_DELAY_CONE,
    HIGH_LIMIT := 0, HIGH_DELAY := T#0s);
  CEL_FV103_TV02_CMD := fv103_cone.VALVE;
  CEL_FV103_TT02_ALM_DEVIATION := fv103_cone.ALM_DEV;

  fv103_press(PV := CEL_FV103_PT01_PV,
    HIGH_LIMIT := PRESS_HIGH_LIMIT, HIGH_DELAY := PRESS_HIGH_DELAY,
    LOW_LIMIT := PRESS_LOW_LIMIT, LOW_DELAY := PRESS_LOW_DELAY);
  CEL_FV103_PT01_ALM_HIGH := fv103_press.ALM_HIGH;
  CEL_FV103_PT01_ALM_LOW := fv103_press.ALM_LOW;

  (* Spunding setpoint to the RIO, absolute psia x 100, every scan. *)
  CEL_FV103_PCV01_SP := spund_fv103_psig + AMBIENT_PSIA;

  (* FV-104 *)
  fv104_side(PV := CEL_FV104_TT01_PV, SP := CEL_FV104_TT01_SP,
    DEV_LIMIT := TEMP_DEV_LIMIT, DEV_DELAY := TEMP_DEV_DELAY_SIDE,
    HIGH_LIMIT := TEMP_HIGH_LIMIT, HIGH_DELAY := TEMP_HIGH_DELAY);
  CEL_FV104_TV01_CMD := fv104_side.VALVE;
  CEL_FV104_TT01_ALM_DEVIATION := fv104_side.ALM_DEV;
  CEL_FV104_TT01_ALM_HIGH := fv104_side.ALM_HIGH;

  fv104_cone(PV := CEL_FV104_TT02_PV, SP := CEL_FV104_TT02_SP,
    DEV_LIMIT := TEMP_DEV_LIMIT, DEV_DELAY := TEMP_DEV_DELAY_CONE,
    HIGH_LIMIT := 0, HIGH_DELAY := T#0s);
  CEL_FV104_TV02_CMD := fv104_cone.VALVE;
  CEL_FV104_TT02_ALM_DEVIATION := fv104_cone.ALM_DEV;

  fv104_press(PV := CEL_FV104_PT01_PV,
    HIGH_LIMIT := PRESS_HIGH_LIMIT, HIGH_DELAY := PRESS_HIGH_DELAY,
    LOW_LIMIT := PRESS_LOW_LIMIT, LOW_DELAY := PRESS_LOW_DELAY);
  CEL_FV104_PT01_ALM_HIGH := fv104_press.ALM_HIGH;
  CEL_FV104_PT01_ALM_LOW := fv104_press.ALM_LOW;

  (* Spunding setpoint to the RIO, absolute psia x 100, every scan. *)
  CEL_FV104_PCV01_SP := spund_fv104_psig + AMBIENT_PSIA;
END_PROGRAM
